RoboDK station: EliteRobotsCS63.rdk

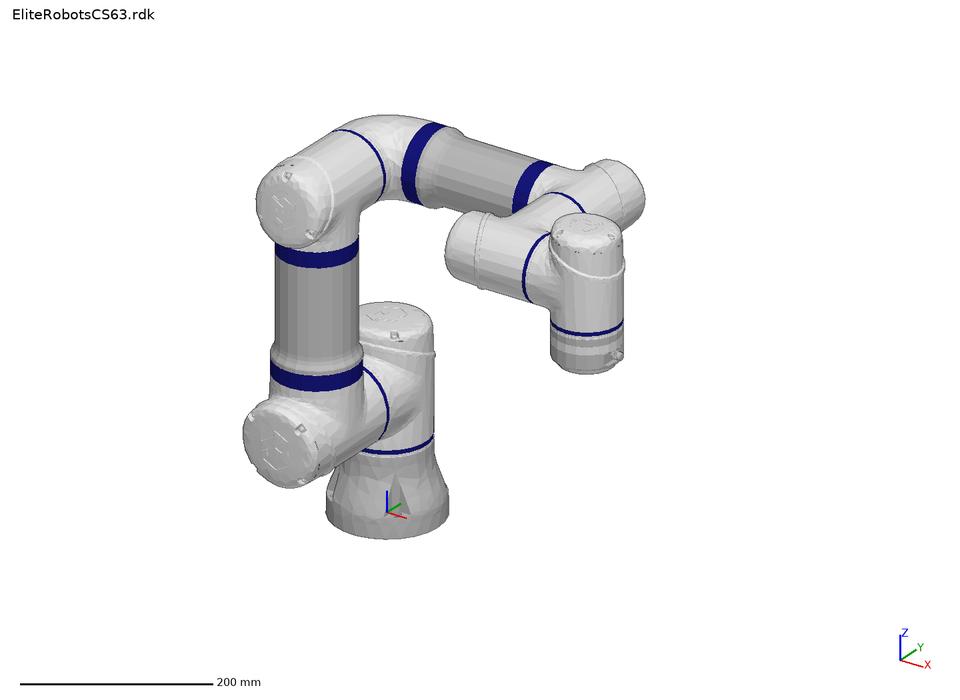
[picture v0: the station drawn from its stored meshes, robots at their saved joint values, targets as dots, program paths as lines]
Station EliteRobotsCS63 (saved by RoboDK 6.2.0). Poses are relative to the parent item; angles as X-Y-Z fixed-axis rotations.
  - frame Elite Robots CS63 Base at (0, 0, 0) mm
    - robot Elite Robots CS63: 6 axes
        modified DH rows (alpha deg, a mm, theta deg, d mm): 0, 0, 0, 153; 90, 0, 180, 0; 0, 270, 0, 0; 0, 257.5, 0, 144.5; -90, 0, 0, 96.5; 90, 0, 180, 92
        joint limits [-360, -360, -360, -360, -360, -360] to [360, 360, 360, 360, 360, 360]; home [0, -90, -90, -90, 90, 0]; saved at [0, -90, -90, -90, 90, 0]
